Fanuc KAREL source: kt00733.KL

-- PROVISIONAL review KL for V770-1; original PC SHA256 8e1d2d7150baead9634ee7752968ff2d0ac7a3ef86bdf80b915ac273e45c8c13
-- Incomplete behavior may be omitted. Consult companion uncertainty JSON. Do not deploy.
PROGRAM KT00733
%NOLOCKGROUP
VAR
  OUT : INTEGER
-- UNRESOLVED_DECL ARG type=002011
BEGIN
  -- UNRESOLVED_PC offsets 5-18; opcodes 22,1D,23
  -- UNRESOLVED_PC offsets 23-27; opcodes 7F
END KT00733
